// TIA Portal V19 export
TYPE "EM05_Output"
   STRUCT
      Status : "EM_Output";
      AgitatorActive : Bool;
      LevelInterlock : Bool;
   END_STRUCT;
END_TYPE
